Yaskawa INFORM job: EMPTY.JBI

/JOB
//NAME EMPTY
//POS
///NPOS 0,0,0,0,0,0
//INST
///DATE 2025/01/01 00:00
///ATTR SC,RW
///GROUP1 RB1,BS1
///GROUP2 ST1
NOP
END
